(* IEC 61131-3 sources: Masterarbeit/sigmatek/lasalclass2/PW022_hardware/Class/SafetyManager (part 2) *)

          // if it has an active connection
          if pHelpManaging^.FlexCon.pFSoEConnection then
            // check if one of the safety number is the list match the one of the managing module
            pHelpHDINT := pPara^.aPara[1]$^HDINT;
            for i := 0 to (pPara^.aPara[0]-1)$UDINT do
              // if the connected number from the HWK is found in the list of connected numbers from the SCP => remember it to send it to the managing module
              if pHelpManaging^.FlexCon.SafetyNumber = pHelpHDINT^ then
                MyPara.aPara[0] := pHelpHDINT^$DINT;

                // stop searching for this managing device
                exit;
              end_if;

              pHelpHDINT += sizeof(HDINT);
            end_for;
          end_if;

          // send the current number for this device
          pHelpManaging^.pThis^.NewInst(#MyPara, #MyResult);

          pHelpManaging := pHelpManaging^.pNext;
        end_while;
      end_if;

//**********************************************************************************************************************************************************
    CMD_HWC_CONVERT_COMPRESSED_HWPATH:

      //Method is used to search through the configuration for the handed over compressed hw path and returns the respective uncompressed hw path

      //pPara^.aPara[0] .. version
      //pPara^.aPara[1] .. comp hw path
      //pPara^.aPara[2] .. comp hw path length
      //pPara^.aPara[3] .. pointer to buffer where hw path will be copied
      //pPara^.aPara[4] .. size of buffer where data will be copied

      //pResult^.aData[0]$DINT .. version
      //pResult^.aData[4]$DINT .. retcode when error (negative) or amount of bytes of hw path

      //Check for valid pointer and data lengths
      if (pPara^.aPara[1] = NIL)
       | (pPara^.aPara[2] = 0)
       | (pPara^.aPara[3] = NIL)
       | (pPara^.aPara[4] = 0) then

        ret_code := ERROR;
        pResult^.uiLng := 8;
        pResult^.aData[0]$DINT := 1;  //version of command
        pResult^.aData[4]$DINT := -1; //Invalid pointer or length
        return;
      end_if;

      if pConfigs = NIL  then
        ret_code := ERROR;
        pResult^.uiLng := 8;
        pResult^.aData[0]$DINT := 1;  //version of command
        pResult^.aData[4]$DINT := -2; //no configs yet
        return;
      end_if;

      pHelpConfigs := pConfigs;

      while pHelpConfigs do

        //Go through module configs
        //=============================================================================================================
        if pHelpConfigs^.pFirstModuleCfg then
          pHelpModuleConf := pHelpConfigs^.pFirstModuleCfg;

          while pHelpModuleConf do

            //Check if we got a valid path and len
            if pHelpModuleConf^.ModuleInfo.pCompPath & pHelpModuleConf^.ModuleInfo.CompPathLen then

              //Check if we found the passed path
              if _memcmp(ptr1:=pPara^.aPara[1]$^void, ptr2:=pHelpModuleConf^.ModuleInfo.pCompPath, cntr:=pPara^.aPara[2]$UDINT) = 0 then

                //we found the compressed hw path, return pointer to normal hw path
                if pPara^.aPara[4] > pHelpModuleConf^.ModuleInfo.PathLen then

                  //Copy path to user pointer
                  _memcpy(ptr1:=pPara^.aPara[3]$^void, ptr2:=pHelpModuleConf^.ModuleInfo.pPath, cntr:=pHelpModuleConf^.ModuleInfo.PathLen);

                  ret_code := READY;
                  pResult^.uiLng := 8;

                  pResult^.aData[0]$DINT := 1;  //version
                  pResult^.aData[4]$DINT := pHelpModuleConf^.ModuleInfo.PathLen;
                  return;

                else
                  ret_code := ERROR;
                  pResult^.uiLng := 8;
                  pResult^.aData[0]$DINT := 1;   //version
                  pResult^.aData[4]$DINT := -3;  //not enough space to copy path
                  return;

                end_if;

              end_if;
            end_if;
            pHelpModuleConf := pHelpModuleConf^.pNext;
          end_while;
        end_if;

        //Go through slave config
        //=============================================================================================================
        if pHelpConfigs^.pFirstSlaveCfg then

          pHelpSlaveCfg := pHelpConfigs^.pFirstSlaveCfg;

          while pHelpSlaveCfg do

            //Check if we got a valid path and len
            if pHelpSlaveCfg^.SlaveInfo.pCompPath & pHelpSlaveCfg^.SlaveInfo.CompPathLen then

              //Check if we found the passed path
              if _memcmp(ptr1:=pPara^.aPara[1]$^void, ptr2:=pHelpSlaveCfg^.SlaveInfo.pCompPath, cntr:=pPara^.aPara[2]$UDINT) = 0 then

                //we found the compressed hw path, return pointer to normal hw path
                if pPara^.aPara[4] > pHelpSlaveCfg^.SlaveInfo.PathLen then

                  //Copy path to user pointer
                  _memcpy(ptr1:=pPara^.aPara[3]$^void, ptr2:=pHelpSlaveCfg^.SlaveInfo.pPath, cntr:=pHelpSlaveCfg^.SlaveInfo.PathLen);

                  ret_code := READY;
                  pResult^.uiLng := 8;

                  pResult^.aData[0]$DINT := 1;  //Path was found
                  pResult^.aData[4]$DINT := pHelpSlaveCfg^.SlaveInfo.PathLen;
                  return;

                else
                  ret_code := ERROR;
                  pResult^.uiLng := 8;
                  pResult^.aData[0]$DINT := 1;   //version
                  pResult^.aData[4]$DINT := -3;  //not enough space to copy path
                  return;

                end_if;
              end_if;
            end_if;
            pHelpSlaveCfg := pHelpSlaveCfg^.pNext;
          end_while;
        end_if;

        //Go through fsoe connections
        //=============================================================================================================
        if pHelpConfigs^.pFirstFSoEConnection then
          pHelpFsoeConn := pHelpConfigs^.pFirstFSoEConnection;

          while pHelpFsoeConn do

            //Check if we got a valid path and len
            if pHelpFsoeConn^.pSlavePathComp & pHelpFsoeConn^.SlavePathLen then

              //Check if we found the passed path
              if _memcmp(ptr1:=pPara^.aPara[1]$^void, ptr2:=pHelpFsoeConn^.pSlavePathComp, cntr:=pPara^.aPara[2]$UDINT) = 0 then

                //we found the compressed hw path, return pointer to normal hw path
                if pPara^.aPara[4] > pHelpFsoeConn^.SlavePathLen then

                  //Copy path to user pointer
                  _memcpy(ptr1:=pPara^.aPara[3]$^void, ptr2:=pHelpFsoeConn^.pSlavePath, cntr:=pHelpFsoeConn^.SlavePathLen);

                  ret_code := READY;
                  pResult^.uiLng := 8;

                  pResult^.aData[0]$DINT := 1;  //Path was found
                  pResult^.aData[4]$DINT := pHelpFsoeConn^.SlavePathLen;
                  return;

                else
                  ret_code := ERROR;
                  pResult^.uiLng := 8;
                  pResult^.aData[0]$DINT := 1;   //version
                  pResult^.aData[4]$DINT := -3;  //not enough space to copy path
                  return;
                end_if;
              end_if;

            end_if;
            pHelpFsoeConn := pHelpFsoeConn^.pNext;
          end_while;
        end_if;

        pHelpConfigs := pHelpConfigs^.pNext;
      end_while;

      //comp hw path was not found in config
      ret_code := ERROR;
      pResult^.uiLng := 8;
      pResult^.aData[0]$DINT := 1;   //version
      pResult^.aData[4]$DINT := -4;  //passed path was not found in configuration list

//**********************************************************************************************************************************************************
  else
    bd_LogRtMessagesInCy.InvalidCommandReceived := TRUE;
  END_CASE;

#ifdef SAFETY_DEBUG_LOGGING_ACTIVATED
  if InitSSW <> OldInitSSW then
#ifdef SAFETY_DEBUG_TRACING_ACTIVATED
    LogValue("@DBG (SafetyManager::ClassState::NewInst) InitSSW changed from {0} to {1}", Value:=OldInitSSW, Value2:=InitSSW);
#endif
    LogBuf[ActLogIndex].NewState := InitSSW;
    LogBuf[ActLogIndex].OldState := OldInitSSW;
    LogBuf[ActLogIndex].Command := 0;
    LogBuf[ActLogIndex].TimeSinceLastLog_us := OS_READMICROSEC();
    LogBuf[ActLogIndex].TimeSinceLastLog_us -= TimeStampLastLog_us;
    TimeStampLastLog_us := OS_READMICROSEC();
    if ActLogIndex = (LogBufferSize - 1) then
      ActLogIndex := 0;
    else
      ActLogIndex += 1;
    end_if;
  end_if;
  OldInitSSW := InitSSW;
#endif

  ret_code := READY;

END_FUNCTION

FUNCTION VIRTUAL GLOBAL SafetyManager::CyWork
  VAR_INPUT
    EAX 	: UDINT;
  END_VAR
  VAR_OUTPUT
    state (EAX) 	: UDINT;
  END_VAR
  VAR
    MyPara 	      : CmdStruct;
    MyResult	    : results;
    pHelpSafety   : ^t_SafetyComponent;
    pHelpManaging : ^t_ManagingComponent;
    pModuleInfo   : ^t_ModuleInfo;
    pTempMem      : ^void;
    i             : UDINT;
    Synchron      : BOOL;
    AllReady      : BOOL;
    pHelpCfg      : ^t_LocalCfgListElem;
    pHelpConfig   : ^t_CfgListElem;
  END_VAR

//=================================================================================================
#ifdef VM_CLASS_TIME_MEASUREMENT
  StartTimeMeasurement(VARANTIME_CY);
#endif
//=================================================================================================
  // if we got UDP stuff going on => start the udp task
  if (sUdpVars.UdpTaskStarted = FALSE) & (sUdpVars.ProducerConnectionNo | ((sUdpVars.UdpInit AND 2#11) = (t_UdpInit.FSoEAvailable OR t_UdpInit.ProvidesIF))) then
    To_MultiTask.CREATETHREAD(taskfunction0 := #UdpTask()
                            , priority0     := 14           // same priority as cyclic task
                            , stackSize0    := 0x4000
                            , flags0        := MT_TASK_SAVETHIS
                            , parameter0    := THIS
                            , name0         := "SafetyUDP");

    sUdpVars.UdpTaskStarted := TRUE;
  end_if;

  case InitSSW of
//**********************************************************************************************************************************************************
    _NotMaster: // don't start any actions, because we're not the master. but if the master wants something from us, we help out

//**********************************************************************************************************************************************************
    _ClearRoutingInfos: // initialize the structures or clean up an old configuration
      if ClearRoutingInformations() then

        // reactivate the domain synchronicity timeout
        b_SynchroTimeoutSet := FALSE;

        InitSSW := _FirstWait4SynchronManagingNodes;
      end_if;

//**********************************************************************************************************************************************************
    _FirstWait4SynchronManagingNodes: // wait for managing nodes to be syncron (all nodes are optionaly for this case, the will be checked later again)
      if SafetyDomainTimeout & (b_SynchroTimeoutSet = FALSE) then
        b_SynchroTimeoutSet := TRUE;
        SynchroTimeout := ops.tAbsolute;
      end_if;

      Synchron := AllManagingNodesSynchron();
                                                        // we wait synchro timeout + 50ms (50ms time for the domains to give up trying: see AllManagingNodesSynchron method)
      if Synchron then// | (SafetyDomainTimeout & ((ops.tAbsolute - SynchroTimeout) > (SafetyDomainTimeout + 50))) then
        if b_SyncTimeoutExceeded then
          b_SyncTimeoutExceeded := FALSE;
          LogError("@0444 (SafetyManager::CyWork) Timeout for managing module (VBC, VMC,..) exceeded! Initialisation will continue to check if it's optional!");
        end_if;

        InitSSW := _SetConnectionOk;
      end_if;

//**********************************************************************************************************************************************************
    _SetConnectionOk:
      // send hw-connection ok to start SDOs
      MyPara.uiCmd := CMD_SM_FIRST_CONNECT_READY;
      MyPara.aPara[0] := 0; // length of parameters

      TellAllSafetyModules(#MyPara, #MyResult);

      b_MandatoryStuffAvailable := FALSE;
      LastCfgReceiveTime := ops.tAbsolute;

      InitSSW := _Wait4ReInit;

//**********************************************************************************************************************************************************
    _Wait4ReInit: // wait until all local CSCPs have a valid configuration before we wait to be synchron with other domains

      // add our local configurations if there are any
      SendLocalCfgsToMaster();

      // wait until we got a valid config of every local safety cpu
      if (LocalCPUCfgNo = LocalCPUNo) | b_MandatoryStuffAvailable then
        AllReady := TRUE;

        if LocalCPUCfgNo then
          pHelpCfg := pFirstLocalCPUCfg;

          // for is used to ensure thread safety
          for i := 0 to (LocalCPUCfgNo-1) do
            if pHelpCfg^.ConfigSize = 0 then
              AllReady := FALSE;
              exit;
            end_if;

            pHelpCfg := pHelpCfg^.pNext;
          end_for;
        end_if;

        // if we have a config from every cscp, we start the initialisation
        if AllReady then
          InitSSW := _CheckLocalCPUConfigs;
        end_if;
      else
        // if we already got a config => check if there is something optional
        if LocalCPUCfgNo & ((ops.tAbsolute - LastCfgReceiveTime) > 5000) then
          CheckOptional();
        end_if;

        InitSSW := _SendInterfaceConfigs;
      end_if;

//**********************************************************************************************************************************************************
    _CheckLocalCPUConfigs: // check for unused and optional modules in the local configurations (needed for correct time synchronisation)
      // if we have a configuration of every safety cpu => check if the managing modules are optional or any of the safety/managing components is unused (not involved in any PDO)
      if (LocalCPUCfgNo = LocalCPUNo) | b_MandatoryStuffAvailable then

        // set the IsOptional-Bit of all modules (safety and managing components) to TRUE
        // in CheckModuleUsage the the non-optional will get the IsOptional-Bit set to FALSE
        pHelpSafety := pFirstSafetyComponent;
        while pHelpSafety do
          pHelpSafety^.InfoBits.IsOptional    := TRUE;

          pHelpSafety := pHelpSafety^.pNext;
        end_while;

        pHelpManaging := pFirstManagingInterfaceComponent;
        while pHelpManaging do
          pHelpManaging^.InfoBits.IsOptional    := TRUE;

          pHelpManaging := pHelpManaging^.pNext;
        end_while;

        // check all configurations which modules are used
        if LocalCPUCfgNo then
          pHelpCfg := pFirstLocalCPUCfg;

          for i := 0 to (LocalCPUCfgNo-1) do
            // check for used modules and mark them in the infobits
            CheckModuleUsage(pHelpCfg^.ConfigSize, pHelpCfg^.pConfig, pHelpCfg^.IsFSoECfg);

            pHelpCfg := pHelpCfg^.pNext;
          end_for;
        end_if;

        // now create the linked list for the time synchronisation
        CreateTimeSyncList();

        if (pFirstManagingInterfaceComponent = NIL) then
          // if we have FSoE Modules => check the connection between the modules and tell them what to copy
          if b_GotFSoEModules then
            CreateFSoEPDOs();

            if b_AllLocalSlaveAddressesValid then
              InitSSW := _NoDomains;
            else
              // wait for all local connections to be established
              SetTimeout();
              InitSSW := _Wait4FSoEConnectionsLocal;
            end_if;
          else
            InitSSW := _NoDomains;
          end_if;
        else
          // reactivate the domain synchronicity timeout, because now we know what is really optional
          b_SynchroTimeoutSet := FALSE;

          InitSSW := _Wait4SynchronManagingNodes;
        end_if;

      end_if;

//**********************************************************************************************************************************************************
    _Wait4FSoEConnectionsLocal:
      CheckTimeout();
      if b_AllLocalSlaveAddressesValid then
        CreateFSoEPDOs();
        // success => continue
        InitSSW := _NoDomains;
      end_if;

//**********************************************************************************************************************************************************
    _Wait4SynchronManagingNodes: // wait until all managing modules are synchron with the other stations
      if SafetyDomainTimeout & (b_SynchroTimeoutSet = FALSE) then
        b_SynchroTimeoutSet := TRUE;
        SynchroTimeout := ops.tAbsolute;
      end_if;

      Synchron := AllManagingNodesSynchron();
                                                        // we wait synchro timeout + 50ms (50ms time for the domains to give up trying: see AllManagingNodesSynchron method)
      if Synchron then// | (SafetyDomainTimeout & ((ops.tAbsolute - SynchroTimeout) > (SafetyDomainTimeout + 50))) then
        if b_SyncTimeoutExceeded then
          b_SyncTimeoutExceeded := FALSE;
          LogError("@0445 (SafetyManager::CyWork) Timeout for optional managing module (VBC, VMC,..) exceeded! Initialisation will continue without it!");
        end_if;

        // add our own safety cpus to the config list
        AddOwnCPUsToList();

        if NewTimeSyncPossible() then
          // tell every safety module, that it has to initialize the memory for writing the time synchronisation
          SetNewSyncMode(TRUE);
          MyPara.aPara[3] := 1;
        else
          SetNewSyncMode(FALSE);
          MyPara.aPara[3] := 0;
        end_if;

        InitSSW := _SendDomainNr;
      end_if;

//**********************************************************************************************************************************************************
    _SendDomainNr: // send the domain nr. to the managing nodes
      // if we have a valid domain number
      MyPara.uiCmd := CMD_SM_DOMAIN_NR_SEND;
      MyPara.aPara[0] := 1; // length of parameters

      pTempMem := NIL;

      if us_SafetyModuleNo then
        if ud_SizeTempMemCy >= 1 + us_SafetyModuleNo * sizeof(t_ModuleInfo) then
          pTempMem := pTempMemCy;
        else
          LogError("@0446 (SafetyManager::CyWork) _SendDomainNr: Temporary memory for cyclic task is too small!");
          LogValue("AvaliableMem: {0} / NeededMem: {1}", Value:=ud_SizeTempMemCy, Value2:=1 + us_SafetyModuleNo * sizeof(t_ModuleInfo));
        end_if;

        if pTempMem then
          MyPara.aPara[1] := pTempMem$DINT;
          pModuleInfo$^void := pTempMem;

          pModuleInfo^$USINT := 0;
          pModuleInfo += sizeof(USINT);
          if pFirstSafetyComponent then
            pHelpSafety := pFirstSafetyComponent;
            while pHelpSafety do
              pModuleInfo^.SafetyNbr := pHelpSafety^.SafetyNbr;

              pHelpSafety := pHelpSafety^.pNext;
              pModuleInfo += sizeof(t_ModuleInfo);
            end_while;

            MyPara.aPara[0] += us_SafetyModuleNo * sizeof(t_ModuleInfo);
          end_if;
        else
          MyPara.aPara[1] := (#MyPara.aPara[3])$DINT;
          MyPara.aPara[3] := 0;
          LogError("@0447 (SafetyManager::CyWork) Failed to allocate memory for distributing the local module information");
        end_if;
      else
        MyPara.aPara[1] := (#MyPara.aPara[3])$DINT;
        MyPara.aPara[3] := 0;
      end_if;

      // tell all interface modules, because maybe they don't know we're an interface neighbor
      TellAllInterfaceManagingModules(#MyPara, #MyResult);

      DomainInfoSendTime := ops.tAbsolute;

      // the slaves get this via newinst command
      InitSSW := _Wait4DomainInfos;

//**********************************************************************************************************************************************************
    _Wait4DomainInfos:
      // wait a little for further domain infos (which are sent as response to our message)
      if (ops.tAbsolute - DomainInfoSendTime) > 200 then
        InitSSW := _Wait4CPUConfigs;
        SetTimeout();
      end_if;

//**********************************************************************************************************************************************************
    _Wait4CPUConfigs:
      CheckTimeout();
      if AllCPUConfigsArrived() then
        // if all needed modules are available (all non-optional modules or interface frames)
        if CheckCPUConfigs() then
          // check if there are PDO configs to broadcast
          if ActPDO_ID then
            // before we broadcast the PDOs, we check if the length informations are correct on every entry
            PDOLengthCorrection();

            // if we have interface-connections, we wait for the safety numbers of it
            if pFirstManagingInterfaceComponent & AnyIFDomainSynchron() then
              InitSSW := _SendInterfaceConfigs;
            else
              InitSSW := _SendNextPDO;
            end_if;
          else
            if pFirstManagingInterfaceComponent & b_GotFSoEModules then
              // we have some FSoE Connections
              InitSSW := _SendInterfaceConfigs;
            else
              // otherwise => finalize initialisation
              InitSSW := _Wait4CopyCmdStart;
            end_if;
          end_if;
        else
          // if configs are not ok => set everything to finished so that the firmware can show the error information (otherwise the firmware will not start doing anything)
          InitSSW := _Wait4CopyCmdStart;
        end_if;
      end_if;

//**********************************************************************************************************************************************************
    _SendInterfaceConfigs:
      // if all domain managing modules needed for non-optional pdos are synchron
      if AllNonOptionalIFDomainsSynchron() then
        if b_GotFSoEModules then
          CreateFSoEPDOs();
        end_if;

        // send our configs to all inferface domains
        SendInterfaceConfigs(NIL, FALSE, b_GotFSoEModules);

        InitSSW := _Wait4InterfaceConfigs;
        SetTimeout();
      end_if;

//**********************************************************************************************************************************************************
    _Wait4InterfaceConfigs:
      CheckTimeout();
      if AllInterfaceCfgsArrived() then
        if (LocalCPUCfgNo = LocalCPUNo) | b_MandatoryStuffAvailable then
          if pActualSendPDO then
            InitSSW := _SendNextPDO;
          else
            if b_GotFSoEModules then
              SetTimeout();
              InitSSW := _Wait4FSoEConnectionsExternal;
            else
              InitSSW := _Wait4ReInit;
            end_if;
          end_if;
        else
          InitSSW := _Wait4ReInit;
        end_If;
      end_if;

//**********************************************************************************************************************************************************
    _Wait4FSoEConnectionsExternal:
      CheckTimeout();
      if b_AllLocalSlaveAddressesValid then
        CreateFSoEPDOs();
        FinalizePDOMapping();
        InitSSW := _FinishInitialisation;
      end_if;

//**********************************************************************************************************************************************************
    _SendNextPDO:
      // broadcast the PDO
      BroadCastActPDO();

      InitSSW := _Wait4PDOAcks;
      SetTimeout();

//**********************************************************************************************************************************************************
    _Wait4PDOAcks:
      // wait until all acknowledges arrive (all modules which are needed for PDO transport have to answer!)
      CheckTimeout();

      // check if there is another PDO configuration to send
      repeat
        if pActualSendPDO^.pNext then
          pActualSendPDO := pActualSendPDO^.pNext;
        else
          if pActualSendCfg^.pNext then
            pActualSendCfg := pActualSendCfg^.pNext;
            pActualSendPDO := pActualSendCfg^.pFirstPdoCfg;

            // if there is no pdo config in this config, go to the next config
            while (pActualSendPDO = NIL) & pActualSendCfg^.pNext do
              pActualSendCfg := pActualSendCfg^.pNext;
              pActualSendPDO := pActualSendCfg^.pFirstPdoCfg;
            end_while;
          else
            pActualSendCfg := NIL;
            pActualSendPDO := NIL;
          end_if;
        end_if;

      // skip double entries
      until ((pActualSendPDO = NIL) | (pActualSendPDO^.PdoInfo.Info.DoublePDOEntry = FALSE)) end_repeat;

      // if we found another PDO => send it
      if pActualSendPDO then
        InitSSW := _SendNextPDO;
      else
        // otherwise => finalize initialisation
        InitSSW := _Wait4CopyCmdStart;
      end_if;

//**********************************************************************************************************************************************************
    _Wait4CopyCmdStart:
      // this step is handlet in RT because the DOs are isochronous

//**********************************************************************************************************************************************************
    _NoDomains:
      // No domains available => just check if there are old modules or new modules used
      if NewTimeSyncPossible() then
        // tell every safety module, that it has to initialize the memory for writing the time synchronisation
        SetNewSyncMode(TRUE);
      else
        SetNewSyncMode(FALSE);
      end_if;

      // we may have internal interface frames and therefore we have to create a list with the local CRCs
      if LocalIFsAvailable() then
        // add local IFs for easier SDO/TDO forwarding
        CheckCPUConfigs();

        // check if there are PDO configs to broadcast
        if ActPDO_ID & (b_GotFSoEModules = FALSE) then
          // before we broadcast the PDOs, we check if the length informations are correct on every entry
          PDOLengthCorrection();

          // distribute PDOs locally
          pHelpConfig := pConfigs;
          while pHelpConfig do
            pActualSendCfg := pHelpConfig;
            pActualSendPDO := pHelpConfig^.pFirstPdoCfg;
            while pActualSendPDO do
              BroadCastActPDO();

              pActualSendPDO := pActualSendPDO^.pNext;
            end_while;

            pHelpConfig := pHelpConfig^.pNext;
          end_while;
        end_if;
      end_if;

      InitSSW := _FinishInitialisation;

//**********************************************************************************************************************************************************
    _FinishInitialisation:
      // if it's the new mode also start the sync process at the first safety device
      MyPara.uiCmd := CMD_SM_INIT_FINISHED;
      MyPara.aPara[0] := 0; // length of parameters

      // sent set bus ready signal (quit error 199 if active)
      TellAllSafetyModules(#MyPara, #MyResult);

      // if we have the new sync mode => start the time synchronisation here
      if b_NewSyncMode then
        b_StartTimeSync := TRUE;
      end_if;

      MinSyncDuration := 16#7FFFFFFF;

      // if there was an error and we still reached this point, don't conceal the error (except if it's a timeout in this init sequence or a SDO problem which could have been fixed)
      if (ClassState = 0) | (ClassState = -11) | (ClassState = -8) then
        ClassState := 1;
      end_if;

      InitSSW := _InitFinished;

//**********************************************************************************************************************************************************
    _InitFinished: // finished with initialisation, now start our cyclic business

      // check sync timeout counter
      if SyncTimeoutCounter >= TIMESYNC_TIMEOUTS_BEFORE_LOGMSG then
        LogError("@0448 (SafetyManager::CyWork) Timeout while Timesynchronizing");

        // reset counter
        SyncTimeoutCounter := 0;
      end_if;

      // print log messages from realtime here to prevent rt-runtime errors
      if bd_LogRtMessagesInCy then
        if bd_LogRtMessagesInCy.NoTDOTargetToManager then
          bd_LogRtMessagesInCy.NoTDOTargetToManager := FALSE;
          LogError("@0449 (SafetyManager::ClassState::NewInst) Couldn't find target of TDO on the way to the manager");
        end_if;

        if bd_LogRtMessagesInCy.NoTDOTargetToModule then
          bd_LogRtMessagesInCy.NoTDOTargetToModule := FALSE;
          LogError("@044A (SafetyManager::ClassState::NewInst) Couldn't find target of TDO on the way to the module");
        end_if;

        if bd_LogRtMessagesInCy.InvalidCommandReceived then
          bd_LogRtMessagesInCy.InvalidCommandReceived := FALSE;
          LogError("@044B (SafetyManager::State::NewInst) Invalid command received");
        end_if;

        if bd_LogRtMessagesInCy.UnkownCopySource then
          bd_LogRtMessagesInCy.UnkownCopySource := FALSE;
          LogError("@044D (SafetyManager::RtWork) Could not activate copy command, because source address is unknown (waiting for safety number info)");
        end_if;

        if bd_LogRtMessagesInCy.InvalidIFConfiguration then
          bd_LogRtMessagesInCy.InvalidIFConfiguration := FALSE;
          LogError("@044E (SafetyManager::GiveTokenToNextModule) Only non-synchron interface domains found => need at least one safe CPU!");
        end_if;

        if bd_LogRtMessagesInCy.TooManyOptionalMissing then
          bd_LogRtMessagesInCy.TooManyOptionalMissing := FALSE;
          LogError("@044F (SafetyManager::GiveTokenToNextModule) Too many optional modules missing for a correct time sync cycle");
        end_if;

        if bd_LogRtMessagesInCy.UdpReceivedInvalidCommand then
          bd_LogRtMessagesInCy.UdpReceivedInvalidCommand := FALSE;
          LogError("@0450 (SafetyManager::ReceiveUdpData) Received invalid command via UDP");
        end_if;

        if bd_LogRtMessagesInCy.UdpReceivedInvalidState then
          bd_LogRtMessagesInCy.UdpReceivedInvalidState := FALSE;
          LogError("@0451 (SafetyManager::ReceiveUdpData) Received invalid state via UDP");
        end_if;

        if bd_LogRtMessagesInCy.UdpNoMem4Connections then
          bd_LogRtMessagesInCy.UdpNoMem4Connections := FALSE;
          LogError("@0452 (SafetyManager::AddIpConnection) Can't add udp connection, since the memory is not allocated");
        end_if;
      end_if;
//**********************************************************************************************************************************************************
  end_case;

#ifdef SAFETY_DEBUG_LOGGING_ACTIVATED
  if InitSSW <> OldInitSSW then
#ifdef SAFETY_DEBUG_TRACING_ACTIVATED
    LogValue("@DBG (SafetyManager::CyWork) InitSSW changed from {0} to {1}", Value:=OldInitSSW, Value2:=InitSSW);
#endif
    LogBuf[ActLogIndex].NewState := InitSSW;
    LogBuf[ActLogIndex].OldState := OldInitSSW;
    LogBuf[ActLogIndex].Command := 0;
    LogBuf[ActLogIndex].TimeSinceLastLog_us := OS_READMICROSEC();
    LogBuf[ActLogIndex].TimeSinceLastLog_us -= TimeStampLastLog_us;
    TimeStampLastLog_us := OS_READMICROSEC();
    if ActLogIndex = (LogBufferSize - 1) then
      ActLogIndex := 0;
    else
      ActLogIndex += 1;
    end_if;
  end_if;
  OldInitSSW := InitSSW;
#endif

  state := READY;

//=================================================================================================
#ifdef VM_CLASS_TIME_MEASUREMENT
  StopTimeMeasurement(VARANTIME_CY);
#endif
//=================================================================================================

END_FUNCTION

FUNCTION SafetyManager::AddModule
  VAR_INPUT
    pPara 	: ^CmdStruct;
  END_VAR
  VAR_OUTPUT
    retcode 	: BOOL;
  END_VAR
  VAR
    ModuleType : t_e_ModuleType;
  END_VAR

  retcode := FALSE;

  ModuleType := pPara^.aPara[0]$t_e_ModuleType;

  // we differ between real safety components and managing components
  case ModuleType of
    _CSCP01x,
    _CSDI16x,
    _CSTO08x,
    _SCP010,
    _SCP011,
    _SCP111,
    _SCP211,
    _MS011,
    _MS012,
    _SDD1300,
    _SDD1400,
    _SDD1500,
    _SDD1600,
    _ModuleWithoutConfig:
        retcode := AddSafetyModule(ModuleType, pPara^.aPara[1]$pVirtualBase);

        if IsFSoEModule(ModuleType) then

          //only allocate memory if it is not done before
          if sUdpVars.pTempSendBufferCy = NIL then
            // allocate memory for the temporary cyclic send buffer
            sUdpVars.pTempSendBufferCy$pVoid := To_StdLib.Malloc(size:=sizeof(t_UdpPacketV2));

            if sUdpVars.pTempSendBufferCy then
              _memset(dest:=sUdpVars.pTempSendBufferCy, usByte:=0, cntr:=sizeof(t_UdpPacketV2));
            else
              SetError(bError:=TRUE, ErrorMessage:=_NO_MEMORY_SENDBUFFER_UDP_ERROR, dError:=0);
              LogError("@0453 (SafetyManager::AddModule) Failed to allocate memory for udp send buffer");
            end_if;
          end_if;

          //only allocate memory if it is not done before
          if sUdpVars.pTempSendBufferIRQ = NIL then
            // allocate memory for the temporary irq send buffer
            sUdpVars.pTempSendBufferIRQ$pVoid := To_StdLib.Malloc(size:=sizeof(t_UdpPacketV2));

            if sUdpVars.pTempSendBufferIRQ then
              _memset(dest:=sUdpVars.pTempSendBufferIRQ, usByte:=0, cntr:=sizeof(t_UdpPacketV2));
            else
              SetError(bError:=TRUE, ErrorMessage:=_NO_MEMORY_SENDBUFFER_UDP_ERROR, dError:=0);
              LogError("@0453 (SafetyManager::AddModule) Failed to allocate memory for udp send buffer");
            end_if;
          end_if;

          //only allocate memory if it is not done before
          if sUdpVars.paConnectionsToProducers = NIL then
            sUdpVars.paConnectionsToProducers$pVoid := To_StdLib.Malloc(size:=sizeof(t_aUdpConnections));

            if sUdpVars.paConnectionsToProducers then
              _memset(dest:=sUdpVars.paConnectionsToProducers, usByte:=0, cntr:=sizeof(t_aUdpConnections));
            else
              SetError(bError:=TRUE, ErrorMessage:=_NO_MEMORY_CONNECTION_BUFFER_UDP_ERROR, dError:=0);
              LogError("@0454 (SafetyManager::AddModule) Failed to allocate memory for udp receive buffer");
            end_if;
          end_if;

          //only allocate memory if it is not done before
          if sUdpVars.paConnectionsToConsumers = NIL then
            sUdpVars.paConnectionsToConsumers$pVoid := To_StdLib.Malloc(size:=sizeof(t_aUdpConnections));

            if sUdpVars.paConnectionsToConsumers then
              _memset(dest:=sUdpVars.paConnectionsToConsumers, usByte:=0, cntr:=sizeof(t_aUdpConnections));
            else
              SetError(bError:=TRUE, ErrorMessage:=_NO_MEMORY_CONNECTION_BUFFER_UDP_ERROR, dError:=0);
              LogError("@0454 (SafetyManager::AddModule) Failed to allocate memory for udp receive buffer");
            end_if;
          end_if;
        end_if;

    _VBC021Master,
    _VBC021Slave, // (is limited to 1 per system, because the system can't sync to different systems at the same time)
    _VMC052,
    _VaranManager4VMC, // VaranManager (VMC052 counterpart is also limited to 1 per system, because the system can't sync to different systems at the same time)
    _GenericTimeSyncMaster,
    _GenericTimeSyncSlave,
    _GenericFSoE:
        retcode := AddManagingModule(ModuleType, pPara^.aPara[1]$pVirtualBase, pPara^.aPara[2]$^USINT);
    _GenericDynamicFSoE:
        retcode := AddGenericDynamic(ModuleType, pPara^.aPara[1]$pVirtualBase, pPara^.aPara[2]$^USINT);
  else
    // invalid module type
    ClassState := -7;
    LogError("@0455 (SafetyManager::AddModule) Invalid ModuleType");
  end_case;

  if retcode then
    LoginCnt += 1;
  end_if;

END_FUNCTION

FUNCTION SafetyManager::AddSafetyModule
  VAR_INPUT
    ModuleType 	: t_e_ModuleType;
    pThis 	: pVirtualBase;
  END_VAR
  VAR_OUTPUT
    retcode 	: BOOL;
  END_VAR
  VAR
    pHelpSafety : ^t_SafetyComponent;
  END_VAR

  if pFirstSafetyComponent = NIL then
    pFirstSafetyComponent$pVoid := To_StdLib.Malloc(size:=sizeof(t_SafetyComponent));
    pHelpSafety := pFirstSafetyComponent;
  else
    pHelpSafety := pFirstSafetyComponent;
    while pHelpSafety^.pNext <> NIL do
      pHelpSafety := pHelpSafety^.pNext;
    end_while;
    pHelpSafety^.pNext$pVoid := To_StdLib.Malloc(size:=sizeof(t_SafetyComponent));
    pHelpSafety := pHelpSafety^.pNext;
  end_if;

  if pHelpSafety <> NIL then
    _memset(dest:=pHelpSafety, usByte:=0, cntr:=sizeof(t_SafetyComponent));
    pHelpSafety^.ModuleType   := ModuleType;
    pHelpSafety^.pThis        := pThis;

//    pHelpSafety^.pNext        := NIL;  // not necessary because of memset

    case ModuleType of
//**********************************************************************************************************************************************************
      _CSCP01x,
      _SCP010,
      _SCP011,
      _SCP111,
      _SCP211,
      _SDD1300,
      _SDD1400,
      _SDD1500,
      _SDD1600:
        LocalCPUNo += 1;

//**********************************************************************************************************************************************************
      _CSDI16x,
      _MS011,
      _MS012:
        pHelpSafety^.InfoBits.OnlyInputs := TRUE;
//**********************************************************************************************************************************************************
    end_case;

    us_SafetyModuleNo += 1;

    retcode := TRUE;
  else
    ClassState := -1;

    retcode := FALSE;
  end_if;

END_FUNCTION

FUNCTION SafetyManager::AddManagingModule
  VAR_INPUT
    ModuleType 	: t_e_ModuleType;
    pThis 	: pVirtualBase;
    pObjectPath 	: ^USINT;
  END_VAR
  VAR_OUTPUT
    retcode 	: BOOL;
  END_VAR
  VAR
    pHelpManaging : ^t_ManagingComponent;
    pMyPath : ^USINT;
  END_VAR

  if pFirstManagingInterfaceComponent = NIL then
    pFirstManagingInterfaceComponent$pVoid := To_StdLib.Malloc(size:=sizeof(t_ManagingComponent));
    pHelpManaging := pFirstManagingInterfaceComponent;
  else
    pHelpManaging := pFirstManagingInterfaceComponent;
    while pHelpManaging^.pNext <> NIL do
      pHelpManaging := pHelpManaging^.pNext;
    end_while;
    pHelpManaging^.pNext$pVoid := To_StdLib.Malloc(size:=sizeof(t_ManagingComponent));
    pHelpManaging := pHelpManaging^.pNext;
  end_if;

  if pHelpManaging <> NIL then
    _memset(dest:=pHelpManaging, usByte:=0, cntr:=sizeof(t_ManagingComponent));
    pHelpManaging^.ModuleType     := ModuleType;
    pHelpManaging^.pThis          := pThis;
    pHelpManaging^.DomainNr       := 16#FF;

    if pObjectPath then
      pMyPath$^void := To_StdLib.Malloc(size:=pObjectPath^ + 2);

      // convert 1 byte length info into 2 byte length info
      if pMyPath then
        pMyPath^$UINT := pObjectPath^$USINT;
        To_StdLib.MemCpy(dest:=pMyPath + 2, source:=pObjectPath + 1, size:=pObjectPath^);
      end_if;
    end_if;

    pHelpManaging^.pModulePath := pMyPath;

  //pHelpManaging^.pNext          := NIL;  // not necessary because of memset

    retcode := TRUE;
  else
    ClassState := -1;

    retcode := FALSE;
  end_if;

END_FUNCTION

FUNCTION SafetyManager::AddGenericDynamic
  VAR_INPUT
    ModuleType 	: t_e_ModuleType;
    pThis 	: pVirtualBase;
    pObjectPath 	: ^USINT;
  END_VAR
  VAR_OUTPUT
    retcode 	: BOOL;
  END_VAR
  VAR
    pHelpManaging : ^t_GenericDynamicComponent;
    pMyPath : ^USINT;
  END_VAR

  if pFirstGenericDynamic = NIL then
    pFirstGenericDynamic$pVoid := To_StdLib.Malloc(size:=sizeof(t_GenericDynamicComponent));
    pHelpManaging := pFirstGenericDynamic;
  else
    pHelpManaging := pFirstGenericDynamic;
    while pHelpManaging^.pNext <> NIL do
      pHelpManaging := pHelpManaging^.pNext;
    end_while;
    pHelpManaging^.pNext$pVoid := To_StdLib.Malloc(size:=sizeof(t_GenericDynamicComponent));
    pHelpManaging := pHelpManaging^.pNext;
  end_if;

  if pHelpManaging <> NIL then
    _memset(dest:=pHelpManaging, usByte:=0, cntr:=sizeof(t_GenericDynamicComponent));
    pHelpManaging^.ModuleType     := ModuleType;
    pHelpManaging^.pThis          := pThis;

    if pObjectPath then
      pMyPath$^void := To_StdLib.Malloc(size:=pObjectPath^ + 2);

      // convert 1 byte length info into 2 byte length info
      if pMyPath then
        pMyPath^$UINT := pObjectPath^$USINT;
        To_StdLib.MemCpy(dest:=pMyPath + 2, source:=pObjectPath + 1, size:=pObjectPath^);
      end_if;
    end_if;

    pHelpManaging^.pModulePath := pMyPath;

  //pHelpManaging^.pNext          := NIL;  // not necessary because of memset

    retcode := TRUE;
  else
    ClassState := -1;

    retcode := FALSE;
  end_if;

END_FUNCTION

FUNCTION SafetyManager::AddSafetyNbr
	VAR_INPUT
		pThis 	: pVirtualBase;
		ud_SafetyNbr 	: HDINT;
		FirmwareVersion 	: HDINT;
		FPGAVersion 	: HSINT;
		PathLen 	: USINT;
		pPath 	: ^USINT;
	END_VAR
	VAR_OUTPUT
		retcode 	: BOOL;
	END_VAR
  VAR
    pHelpSafety             : ^t_SafetyComponent;
    pHelpConfigManager      : ^t_CfgListElem;
    pHelpConnectionManager  : ^t_FSoEConnectionDetails;
    pHelpModuleCfg          : ^t_ModuleListElem;
    MyPara 	                : CmdStruct;
    MyResult	              : results;
    pOwnerSafety            : ^t_SafetyComponent;
  END_VAR

  retcode := FALSE;

  if pFirstSafetyComponent then
    pHelpSafety := pFirstSafetyComponent;
    while pHelpSafety do
      if pHelpSafety^.pThis = pThis then
        pHelpSafety^.SafetyNbr    := ud_SafetyNbr;
        pHelpSafety^.FW_Version   := FirmwareVersion;
        pHelpSafety^.FPGA_Version := FPGAVersion;
        pHelpSafety^.PathLen      := PathLen;
        pHelpSafety^.pPath        := pPath;

        if pHelpSafety^.ModuleType = _ModuleWithoutConfig then

          // if the post init is finished => module added during runtime
          if b_PostInitFinished then

            // check all configs
            pHelpConfigManager := pConfigs;
            while pHelpConfigManager do

              // check for FSoE connections that haven't been initialized
              pHelpConnectionManager := pHelpConfigManager^.pFirstFSoEConnection;
              while pHelpConnectionManager do

                if pHelpConnectionManager^.Flags.FSoESlaveHasNoConfig & pHelpConnectionManager^.Flags.IsMaster then
                  if pHelpConnectionManager^.InternalConnectionState = FCS_RESET then
                    ShareSingleConnectionInfos(pHelpConnectionManager, pHelpConfigManager^.pFirstModuleCfg);
                  end_if;
                end_if;

                pHelpConnectionManager := pHelpConnectionManager^.pNext;
              end_while;

              // check all module configs for a match of the path and inform the owner that there is a new safety number
              pHelpModuleCfg := pHelpConfigManager^.pFirstModuleCfg;
              while pHelpModuleCfg do
                if (pHelpModuleCfg^.ModuleInfo.pPath^ = pPath^) &
                   (To_StdLib.MemCmp(pPath + 1, pHelpModuleCfg^.ModuleInfo.pPath + 2 + pHelpModuleCfg^.ModuleInfo.pPath^ - pPath^, pPath^) = 0) then

                  // found a match => tell the owner of the configuration we found the module in

                  pOwnerSafety := pFirstSafetyComponent;
                  while pOwnerSafety do
                    if pOwnerSafety^.SafetyNbr = pHelpConfigManager^.SafetyNbr then
                      MyPara.uiCmd    := CMD_SM_UPDATE_SAFETY_NBR;
                      MyPara.aPara[0] := pHelpModuleCfg^.ModuleInfo.CompPathLen;    // length of HW path
                      MyPara.aPara[1] := pHelpModuleCfg^.ModuleInfo.pCompPath$DINT; // pointer to HW path
                      MyPara.aPara[2] := ud_SafetyNbr$DINT;                         // new safety number
                      pOwnerSafety^.pThis^.NewInst(#MyPara, #MyResult);
                    end_if;

                    pOwnerSafety := pOwnerSafety^.pNext;
                  end_while;
                end_if;

                pHelpModuleCfg := pHelpModuleCfg^.pNext;
              end_while;

              pHelpConfigManager := pHelpConfigManager^.pNext;
            end_while;
          end_if;
        end_if;

        retcode := TRUE;
        return;
      end_if;

      pHelpSafety := pHelpSafety^.pNext;
    end_while;
  end_if;

END_FUNCTION

FUNCTION SafetyManager::GetModuleTypeNo
  VAR_INPUT
    ModuleType 	: t_e_ModuleType;
  END_VAR
  VAR_OUTPUT
    ModuleNo 	: UDINT;
  END_VAR
  VAR
    pHelpSafety   : ^t_SafetyComponent;
    pHelpManaging : ^t_ManagingComponent;
    pHelpGeneric        : ^t_GenericDynamicComponent;
  END_VAR

  ModuleNo := 0;

  if pFirstSafetyComponent then
    pHelpSafety := pFirstSafetyComponent;
    while pHelpSafety do
      if pHelpSafety^.ModuleType = ModuleType then
        ModuleNo += 1;
      end_if;

      pHelpSafety := pHelpSafety^.pNext;
    end_while;
  end_if;

  if pFirstManagingInterfaceComponent then
    pHelpManaging := pFirstManagingInterfaceComponent;
    while pHelpManaging do
      if pHelpManaging^.ModuleType = ModuleType then
        ModuleNo += 1;
      end_if;

      pHelpManaging := pHelpManaging^.pNext;
    end_while;
  end_if;

  if pFirstGenericDynamic then
    pHelpGeneric := pFirstGenericDynamic;

    while pHelpGeneric do
      if pHelpGeneric^.ModuleType = ModuleType then
        ModuleNo += 1;
      end_if;

      pHelpGeneric := pHelpGeneric^.pNext;
    end_while;

  end_if;

END_FUNCTION

FUNCTION SafetyManager::NewTimeSyncPossible
  VAR_OUTPUT
    retcode 	: BOOL;
  END_VAR
  VAR
    pHelpSafety   : ^t_SafetyComponent;
  END_VAR

  // if there is FSoE in the project => no timesync
  if b_GotFSoEModules then
    retcode := FALSE;
    return;
  end_if;

  // default is: we can => check if there is any module with too old firmware or fpga
  retcode := TRUE;

  if pFirstSafetyComponent then
    pHelpSafety := pFirstSafetyComponent;
    while pHelpSafety do

      // check all modules for correct versions
      if ((pHelpSafety^.ModuleType = _CSCP01x) & (   (pHelpSafety^.FPGA_Version    < 16#14)     // if its a CSCP and the FPGA Version is lower than 1.4
                                                   | (pHelpSafety^.FW_Version$UINT < 100)) &    // or the firmware version is lower than 100
                                                      pHelpSafety^.SafetyNbr)                   // only if there is a safety number available (maybe the module is optional and not available)
      |  (pHelpSafety^.NewConfigType = ConfigState_Old) then                                    // or the module has an old config type

        retcode := FALSE;
      end_if;

      pHelpSafety := pHelpSafety^.pNext;
    end_while;
  end_if;

END_FUNCTION

FUNCTION SafetyManager::SetNewSyncMode
  VAR_INPUT
    b_NewMode 	: BOOL;
  END_VAR
  VAR
    MyPara 	  : CmdStruct;
    MyResult	: results;
  END_VAR

  b_NewSyncMode := b_NewMode;

  MyPara.uiCmd := CMD_SM_SET_NEW_SYNC_MODE;
  MyPara.aPara[0] := b_NewSyncMode;
  TellAllSafetyModules(#MyPara, #MyResult);

END_FUNCTION

FUNCTION SafetyManager::TellAllSafetyModules
  VAR_INPUT
    pPara 	: ^CmdStruct;
    pResult 	: ^results;
  END_VAR
  VAR
    pHelpSafety : ^t_SafetyComponent;
  END_VAR

  if pFirstSafetyComponent then
    pHelpSafety := pFirstSafetyComponent;
    while pHelpSafety do
      // call the newinst with the given parameters
      pHelpSafety^.pThis^.NewInst(pPara, pResult);

      pHelpSafety := pHelpSafety^.pNext;
    end_while;
  end_if;

END_FUNCTION

FUNCTION SafetyManager::StartTimeSync

  if pFirstTimeSyncElement then
    pActTimeSyncElement := pFirstTimeSyncElement;

    // send the token to the right module
    GiveTokenToNextModule();

    // remember the start time for calculating the time of a complete synchronisation
    TimeSyncCycleStart := ops.tAbsolute;
  end_if;

END_FUNCTION

FUNCTION SafetyManager::NextTimeSyncModule

  pActTimeSyncElement := pActTimeSyncElement^.pNext;

  // must be done after selecting the new element
  if GiveTokenToNextModule() then
    // we're finished with our synchronisation cycle and just started a new one (must be done after selecting the new element)
    if IsTimeSyncMaster then
      SyncDuration := ops.tAbsolute - TimeSyncCycleStart;
      if SyncDuration > MaxSyncDuration then
        MaxSyncDuration := SyncDuration;
      end_if;
      if SyncDuration < MinSyncDuration then
        MinSyncDuration := SyncDuration;
      end_if;

      // if a cycle has been finished => reset the timeout counter
      SyncTimeoutCounter := 0;

      // remember the start time for calculating the time of a complete synchronisation
      TimeSyncCycleStart := ops.tAbsolute;
    end_if;
  end_if;

END_FUNCTION

FUNCTION SafetyManager::GiveTokenToNextModule
  VAR_OUTPUT
    RestartCycle 	: BOOL;
  END_VAR
  VAR
    MyPara 	  : CmdStruct;
    MyResult	: results;
    pTemp : ^t_TimeSyncElement;
  END_VAR

  if pActTimeSyncElement = pFirstTimeSyncElement then
    RestartCycle := TRUE;
  else
    RestartCycle := FALSE;
  end_if;

  // check if we have to skip something (missing optional modules)
  if TimeSyncModuleAvailable(pActTimeSyncElement) = FALSE then
    // save the actual position
    pTemp := pActTimeSyncElement;

    // if it's a missing optional module
    while (TimeSyncModuleAvailable(pActTimeSyncElement) = FALSE) do
      // skip it
      pActTimeSyncElement := pActTimeSyncElement^.pNext;

      // if we jumped on the first, we have to restart the cycle (time measurement and timeout surveillance)
      if pActTimeSyncElement = pFirstTimeSyncElement then
        RestartCycle := TRUE;
      end_if;

      // if we're at the start of the rotation => stop rotating and print error message
      if pActTimeSyncElement = pTemp then
        bd_LogRtMessagesInCy.TooManyOptionalMissing := TRUE;
        ClassState := -12;
        exit;
      end_if;
    end_while;
  end_if;

  // check if we have to skip something
  if pActTimeSyncElement^.InfoBits.IsInterfaceDomain then
    // save the actual position
    pTemp := pActTimeSyncElement;

    // if it's an interface managing module and it's not synchron, skip it (there has to be also a Safety CPU in the system, therefore we don't ask for it
    while pActTimeSyncElement^.InfoBits.IsInterfaceDomain & (pActTimeSyncElement^.pManaging^.InfoBits.IsSynchron = FALSE) do
      // skip it
      pActTimeSyncElement := pActTimeSyncElement^.pNext;

      // if we jumped on the first, we have to restart the cycle (time measurement and timeout surveillance)
      if pActTimeSyncElement = pFirstTimeSyncElement then
        RestartCycle := TRUE;
      end_if;

      // if we're at the start of the rotation => stop rotating and print error message
      if pActTimeSyncElement = pTemp then
        bd_LogRtMessagesInCy.InvalidIFConfiguration := TRUE;
        ClassState := -12;
        exit;
      end_if;
    end_while;
  end_if;

  if pActTimeSyncElement^.InfoBits.IsConnectionToMaster then
    // don't check for sync timeout if we're not the master
    b_CheckTimeSyncTimeout := FALSE;
  else
    b_CheckTimeSyncTimeout := TRUE;
  end_if;

  // if it's a managing module and not the connection to the master, we give the token to a slave => remember it
  if pActTimeSyncElement^.InfoBits.IsManagingModule & (pActTimeSyncElement^.InfoBits.IsConnectionToMaster = FALSE) then
    b_SlaveSyncActive := TRUE;
  end_if;

  // tell the next module, to start the time synchronisation
  MyPara.uiCmd := CMD_SM_START_TIME_SYNC;
  pActTimeSyncElement^.pThis^.NewInst(#MyPara, #MyResult);

  LastTimeSyncThis := pActTimeSyncElement^.pThis;
  TimeSyncTimeStamp := ops.tAbsolute;

END_FUNCTION

FUNCTION SafetyManager::TellAllInterfaceManagingModules
  VAR_INPUT
    pPara 	: ^CmdStruct;
    pResult 	: ^results;
    OverrideSync 	: BOOL;(* := FALSE *)
  END_VAR
  VAR
    pHelpManaging : ^t_ManagingComponent;
  END_VAR

  if pFirstManagingInterfaceComponent then
    pHelpManaging := pFirstManagingInterfaceComponent;
    while pHelpManaging do
      // call the newinst with the given parameters
      if pHelpManaging^.InfoBits.IsSynchron | OverrideSync then
        pHelpManaging^.pThis^.NewInst(pPara, pResult);
      end_if;

      pHelpManaging := pHelpManaging^.pNext;
    end_while;
  end_if;

END_FUNCTION

FUNCTION SafetyManager::SafetyManager
  VAR_OUTPUT
    ret_code 	: ConfStates;
  END_VAR
  VAR
    sd_retval : DINT;
  END_VAR

  //get interface for hardwaretree functions
  if ( OS_CILGET(INTERFACE_HARDWARETREE, #pHardwareTree)) then
    pHardwareTree := NIL;

    // logging can be used here already because the constructor of the base has been called before to initialize the log-interface-pointer
    LogError("@0457 (SafetyManager::SafetyManager) Hardwaretree-Interface not found. A newer OS is required for Safety-Modules");
  end_if;

  pTempMemCy := To_StdLib.Malloc(size:=SIZE_TEMP_MEMORY);
  if pTempMemCy then
    ud_SizeTempMemCy := SIZE_TEMP_MEMORY;
  else
    LogError("@0458 (SafetyManager::SafetyManager) Allocate temporary Memory failed");
  end_if;

  // try the new interface first
  sd_retval := OS_CILGet(INTERFACE_SAFETY_DLL2, #pSafetyDll2)$DINT;

  if sd_retval then
    // the new safety interface is not available => try the old one
    sd_retval := OS_CILGet(INTERFACE_SAFETY_DLL, #pSafetyDll)$DINT;

    if sd_retval then
      // no dll available
    elsif pSafetyDll^.version >= 5 then
      // dll available that allows quit error
      QuitErrorAvailable := 1;
    end_if;
  else
    // dll available that allows quit error and multiple connections
    QuitErrorAvailable := 2;
  end_if;

  OS_CILGet( INTERFACE_VARANMANAGER, #pVaran );

  ret_code := C_OK;

END_FUNCTION

FUNCTION SafetyManager::AllManagingNodesSynchron
  VAR_OUTPUT
    AllReady 	: BOOL;
  END_VAR
  VAR
    pHelpManaging : ^t_ManagingComponent;
    MyPara 	  : CmdStruct;
    MyResult	: results;
  END_VAR

  AllReady := TRUE;

  // check if any of the managing interface modules is not synchron
  if pFirstManagingInterfaceComponent then
    MyPara.uiCmd := CMD_SM_SYNC_CHECK;

    pHelpManaging := pFirstManagingInterfaceComponent;
    while pHelpManaging do
      // if any managing component isn't synchron => stop searching
      if pHelpManaging^.pThis^.NewInst(#MyPara, #MyResult) = ERROR then
        if (pHelpManaging^.InfoBits.IsOptional = TRUE) then
          if ((SafetyDomainTimeout & ((ops.tAbsolute - SynchroTimeout) > SafetyDomainTimeout))) then
            // we give up waiting => timeout exceeded
            b_SyncTimeoutExceeded := TRUE;
            // if it's the last managing module, then it's our connection to the master module
            if (IsTimeSyncMaster = 0) & pHelpManaging^.InfoBits.IsConnectionToMaster then
              // we have to be our own master now
              IsTimeSyncMaster := 1;
            end_if;
          else
            AllReady := FALSE;
          end_if;
        else
          AllReady := FALSE;
        end_if;

        // return; don't give up here => we have to check it for all domains, this one may be an optional interface frame domain
        pHelpManaging^.InfoBits.IsSynchron := FALSE;
      else
        pHelpManaging^.InfoBits.IsSynchron := TRUE;
      end_if;

      pHelpManaging := pHelpManaging^.pNext;
    end_while;
  end_if;

END_FUNCTION

FUNCTION SafetyManager::GetMasterConnection
  VAR_OUTPUT
    pMasterConn : ^t_ManagingComponent;
  END_VAR
  VAR
    pHelpManaging : ^t_ManagingComponent;
  END_VAR

  pMasterConn := NIL;

  if pFirstManagingInterfaceComponent then
    pHelpManaging := pFirstManagingInterfaceComponent;
    while pHelpManaging do
      if (pHelpManaging^.ModuleType = _VBC021Slave) | (pHelpManaging^.ModuleType = _VaranManager4VMC) | (pHelpManaging^.ModuleType = _GenericTimeSyncSlave) then
        pMasterConn := pHelpManaging;
        pMasterConn^.InfoBits.IsConnectionToMaster := TRUE;
        // if it's not the last in the list => we have to put it in the last place for easier timesync handling (last managing module to handle is the connection back to the master)
        if pMasterConn^.pNext then
          // if it's the first one
          if pMasterConn = pFirstManagingInterfaceComponent then
            pHelpManaging := pFirstManagingInterfaceComponent;
            while pHelpManaging^.pNext do
              pHelpManaging := pHelpManaging^.pNext;
            end_while;
            pFirstManagingInterfaceComponent := pFirstManagingInterfaceComponent^.pNext;
            pHelpManaging^.pNext := pMasterConn;
            pMasterConn^.pNext := NIL;
          else
            // if it's one in the middle
            pHelpManaging := pFirstManagingInterfaceComponent;
            while pHelpManaging^.pNext do
              if pHelpManaging^.pNext = pMasterConn then
                pHelpManaging^.pNext := pMasterConn^.pNext;
              end_if;

              pHelpManaging := pHelpManaging^.pNext;
            end_while;
            pHelpManaging^.pNext := pMasterConn;
            pMasterConn^.pNext := NIL;
          end_if;
        end_if;
        return;
      end_if;

      pHelpManaging := pHelpManaging^.pNext;
    end_while;
  end_if;

END_FUNCTION

FUNCTION SafetyManager::AddConfiguration
  VAR_INPUT
    Length 	: UINT;
    pData 	: ^void;
    IsFSoEConfig 	: BOOL;
  END_VAR
  VAR_OUTPUT
    retcode 	: DINT;
  END_VAR
  VAR
    pHelpCfg          : ^t_CfgListElem;
    pHelpModule       : ^t_ModuleListElem;
    pHelpPdo          : ^t_PdoListElem;
    pHelpSlave        : ^t_SlaveListElem;
    pHelpConnection   : ^t_FSoEConnectionDetails;
    pDataHelp         : ^void;
    i                 : UDINT;
    TmpPathLen        : UINT;
    TempCfgNo         : USINT;
    TempConnectionNo  : UINT;
    pHelpSafety       : ^t_SafetyComponent;
    pHelpManaging     : ^t_ManagingComponent;
    ModuleNo          : UDINT;
  END_VAR

(*
    Memory structure:
      4 Byte: SafetyNumber of CPU (is already there from initialisation in CSCP011_IM::InitSafeModule)
      1 Byte: Number of module configurations which are following
      for every module configuration (first is always the CPU itself)
        1 Byte: Info
        4 Byte: Interface Frame Source SafetyNumber (0 if it is no source for interface frames)
        4 Byte: Interface Frame CRC
        1 Byte: Number of destination inferface frame CRCs
        x Byte: Destination interface frame CRCs (number * sizeof(HDINT)
        2 Byte: Length of hardware path
        x Byte (depending on length in the 2 byte before): Hardwarepath
        2 Byte: Length of compressed hardware path
        x Byte (depending on length in the 2 byte before): Compressed Hardwarepath
        1 Byte: PDO out length for this module
      1 Byte: Number of pdo configurations which are following
      for every PDO configuration
        1 Byte: PDO length
        1 Byte: Interface frame info
        4 Byte: Interface CRC
        2 Byte: Length of source hardware path
        x Byte (depending on length in the 2 byte before): Hardwarepath of source
        2 Byte: Length of destination hardware path
        x Byte (depending on length in the 2 byte before): Hardwarepath of destination
      1 Byte: Number of slave configurations which are following
      for every slave configuration
        1 Byte: Info
        4 Byte: InterfaceCRC
        2 Byte: Length of hardware path
        x Byte (depending on length in the 2 byte before): Hardwarepath
        2 Byte: Length of compressed hardware path
        x Byte (depending on length in the 2 byte before): Compressed Hardwarepath

      if IsFSoEConfig = TRUE
      2 Byte: Number of connection infos which are following
      for every FSoE connection info
        2 Byte: ConnectionID
        1 Byte: ConnectionState
        1 Byte: Flags // Actually, type is 4 bytes in size but for compatibility reasons it is still used as 1 byte. As a result, bits 9-32 are currently not used.
        4 Byte: Master safety number

only if feature available:
        2 Byte: Transmission time in ms

        2 Byte: Offset where to read from master
        2 Byte: Size of data to read from master (and write to slave)
        2 Byte: Offset where to write to master
        2 Byte: Size of data to write to master (and read from slave)
        2 Byte: SlaveAddress
        2 Byte: Length of slave hardware path
        x Byte (depending on length in the 2 byte before): Slave hardware path
        2 Byte: Length of compressed slave hardware path
        x Byte (depending on length in the 2 byte before): Compressed slave hardware path
        2 Byte: Offset where to read from slave
        2 Byte: Offset where to write to slave

*)

  // check if the configuration is valid (pData <> NIL) & (Length must be at least 4 byte for SafetyNbr + 1 byte module cfg number + 1 byte pdo cfg number + 1 byte slave crc number)
  if pData & (Length >= 7)  then

    retcode := 0;

    // first we have to allocate some memory for the configuration
    if pConfigs = NIL then
      pConfigs$pVoid := To_StdLib.Malloc(size:=sizeof(t_CfgListElem));
      pHelpCfg := pConfigs;
    else
      pHelpCfg := pConfigs;
      while pHelpCfg^.pNext <> NIL do
        //if searched path is found, we already got this module in our list
        if pHelpCfg^.SafetyNbr = pData^$HDINT then
          // already in buffer => leave function
          return;
        else
          pHelpCfg := pHelpCfg^.pNext;
        end_if;
      end_while;

      //if searched path is found, we already got this module in our list
      if pHelpCfg^.SafetyNbr = pData^$HDINT then
        // already in buffer => leave function
        return;
      end_if;

      pHelpCfg^.pNext$pvoid := To_StdLib.Malloc(size:=sizeof(t_CfgListElem));
      pHelpCfg := pHelpCfg^.pNext;
    end_if;

    // if we have memory for the configuration => we add the data to the new element
    if pHelpCfg <> NIL then
      pDataHelp := pData;

      // set the next pointer to NIL
      pHelpCfg^.pNext := NIL;

      // safety number of the safety cpu
      pHelpCfg^.SafetyNbr := pDataHelp^$HDINT;
      pDataHelp += sizeof(HDINT);

      // number of module configurations which follow now
      TempCfgNo := pDataHelp^$USINT;
      pDataHelp += sizeof(USINT);

      pHelpCfg^.pFirstModuleCfg := NIL;

      // module configurations
      if TempCfgNo then
        for i := 0 to (TempCfgNo-1) do
          if pHelpCfg^.pFirstModuleCfg = NIL then
            pHelpCfg^.pFirstModuleCfg$pVoid := To_StdLib.Malloc(size:=sizeof(t_ModuleListElem));
            pHelpModule := pHelpCfg^.pFirstModuleCfg;
          else
            pHelpModule^.pNext$pvoid := To_StdLib.Malloc(size:=sizeof(t_ModuleListElem));
            pHelpModule := pHelpModule^.pNext;
          end_if;

          if pHelpModule then
            // initialize the pointers with NIL in case one of the mallocs fails
            pHelpModule^.ModuleInfo.pDestCRCs   := NIL;
            pHelpModule^.ModuleInfo.pPath       := NIL;
            pHelpModule^.ModuleInfo.pCompPath   := NIL;
            pHelpModule^.pNext                  := NIL;

            // info
            pHelpModule^.ModuleInfo.Info := pDataHelp^$BSINT;
            pDataHelp += sizeof(BSINT);

            // safety number of interface frame source
            pHelpModule^.ModuleInfo.SafetyNbr := pDataHelp^$HDINT;
            pDataHelp += sizeof(HDINT);

            // if it's the config owner => take the address service info to the info bits
            if pHelpCfg^.SafetyNbr = pHelpModule^.ModuleInfo.SafetyNbr then
              pHelpSafety := pFirstSafetyComponent;
              while pHelpSafety do
                // check if we got a component with this number
                if pHelpSafety^.SafetyNbr = pHelpCfg^.SafetyNbr then
                  pHelpSafety^.InfoBits.IsAddressService := pHelpModule^.ModuleInfo.Info.IsAddressService;
                end_if;

                pHelpSafety := pHelpSafety^.pNext;
              end_while;
            end_if;

            // interface CRC of interface frame
            pHelpModule^.ModuleInfo.InterfaceCRC := pDataHelp^$HDINT;
            pDataHelp += sizeof(HDINT);

            if pHelpModule^.ModuleInfo.InterfaceCRC then
              // someone might connect to us via udp because we supply an interface frame
              sUdpVars.UdpInit.ProvidesIF := TRUE;
            end_if;

            // interface frame destination CRCs
            if pHelpModule^.ModuleInfo.Info.IsInterfaceDest then
              // number of CRCs
              TmpPathLen := pDataHelp^$USINT; // save some time with this local variable
              pHelpModule^.ModuleInfo.DestCRCNo := TmpPathLen$USINT;
              pDataHelp += sizeof(USINT);

              // allocate memory for the module path
              pHelpModule^.ModuleInfo.pDestCRCs$pVoid := To_StdLib.Malloc(size:=TmpPathLen * sizeof(HDINT));
              if pHelpModule^.ModuleInfo.pDestCRCs = NIL then
                ClassState := -1;
                retcode := -2;
                return;
              end_if;

              // save CRCs
              _memcpy(ptr1:=pHelpModule^.ModuleInfo.pDestCRCs, ptr2:=pDataHelp, cntr:=TmpPathLen * sizeof(HDINT));
              pDataHelp += TmpPathLen * sizeof(HDINT);
            else
              pHelpModule^.ModuleInfo.DestCRCNo := 0;
              pHelpModule^.ModuleInfo.pDestCRCs := NIL;
            end_if;

            // length of hardwarepath
            TmpPathLen := pDataHelp^$UINT; // save some time with this local variable
            pHelpModule^.ModuleInfo.PathLen := TmpPathLen;
            pDataHelp += sizeof(UINT);

            // allocate memory for the module path
            pHelpModule^.ModuleInfo.pPath$pVoid := To_StdLib.Malloc(size:=TmpPathLen);
            if pHelpModule^.ModuleInfo.pPath = NIL then
              ClassState := -1;
              retcode := -2;
              return;
            end_if;

            // save hardwarepath
            _memcpy(ptr1:=pHelpModule^.ModuleInfo.pPath, ptr2:=pDataHelp, cntr:=TmpPathLen);
            pDataHelp += TmpPathLen;

            // length of hardwarepath
            TmpPathLen := pDataHelp^$UINT; // save some time with this local variable
            pHelpModule^.ModuleInfo.CompPathLen := TmpPathLen;
            pDataHelp += sizeof(UINT);

            // allocate memory for the module path
            pHelpModule^.ModuleInfo.pCompPath$pVoid := To_StdLib.Malloc(size:=TmpPathLen);
            if pHelpModule^.ModuleInfo.pCompPath = NIL then
              ClassState := -1;
              retcode := -2;
              return;
            end_if;

            // save compressed hardwarepath
            _memcpy(ptr1:=pHelpModule^.ModuleInfo.pCompPath, ptr2:=pDataHelp, cntr:=TmpPathLen);
            pDataHelp += TmpPathLen;

            // PDO out length for this module (to assign the length to the pdo configurations)
            pHelpModule^.ModuleInfo.PdoOutLen := pDataHelp^$USINT;
            pDataHelp += sizeof(USINT);
          else
            ClassState := -1;
            retcode := -2;
            return;
          end_if;
        end_for;
      end_if;

      // number of Pdo configurations which follow now
      TempCfgNo := pDataHelp^$USINT;
      pDataHelp += sizeof(USINT);

      pHelpCfg^.pFirstPdoCfg := NIL;

      // Pdo configurations
      if TempCfgNo then
        for i := 0 to (TempCfgNo-1) do
          if pHelpCfg^.pFirstPdoCfg = NIL then
            pHelpCfg^.pFirstPdoCfg$pVoid := To_StdLib.Malloc(size:=sizeof(t_PdoListElem));
            pHelpPdo := pHelpCfg^.pFirstPdoCfg;
          else
            pHelpPdo^.pNext$pvoid := To_StdLib.Malloc(size:=sizeof(t_PdoListElem));
            pHelpPdo := pHelpPdo^.pNext;
          end_if;

          if pHelpPdo then
            // initialize the pointers with NIL in case one of the mallocs fails
            pHelpPdo^.PdoInfo.pSourcePath     := NIL;
            pHelpPdo^.PdoInfo.pDestPath       := NIL;
            pHelpPdo^.pNext                   := NIL;

            // pdo length
            pHelpPdo^.PdoInfo.PdoLen := pDataHelp^$USINT;
            pDataHelp += sizeof(USINT);

            // is it an interface pdo?
            pHelpPdo^.PdoInfo.Info := pDataHelp^$BSINT;
            pDataHelp += sizeof(BSINT);

            // if it is an interface frame, we have to copy the CRC too
            if pHelpPdo^.PdoInfo.Info.IsInterfacePDO then
              // interface CRC
              pHelpPdo^.PdoInfo.InterfaceCRC := pDataHelp^$HDINT;
            else
              pHelpPdo^.PdoInfo.InterfaceCRC := 0;
            end_if;
            pDataHelp += sizeof(HDINT);

            // length of source hardwarepath
            TmpPathLen := pDataHelp^$UINT; // save some time with this local variable
            pHelpPdo^.PdoInfo.SourcePathLen := TmpPathLen;
            pDataHelp += sizeof(UINT);

            // allocate memory for the source module path
            pHelpPdo^.PdoInfo.pSourcePath$pVoid := To_StdLib.Malloc(size:=TmpPathLen);
            if pHelpPdo^.PdoInfo.pSourcePath = NIL then
              ClassState := -1;
              retcode := -2;
              return;
            end_if;

            // save source hardwarepath
            _memcpy(ptr1:=pHelpPdo^.PdoInfo.pSourcePath, ptr2:=pDataHelp, cntr:=TmpPathLen);
            pDataHelp += TmpPathLen;

            // check for an IP Address
            if pHelpPdo^.PdoInfo.Info.SrcPathIsCompressed & (pHelpPdo^.PdoInfo.pSourcePath^$USINT = INTERFACE_IP_MODE) then
              // add the connection (we're consumer and we got the IP address of the producer)
              AddUdpConnection(IP:=(pHelpPdo^.PdoInfo.pSourcePath$^HDINT + 5)^, IFCRC:=(pHelpPdo^.PdoInfo.pSourcePath$^HDINT + 1)^, SafetyNumber:=pHelpCfg^.SafetyNbr, ProducerList:=TRUE);
            end_if;

            // length of destination hardwarepath
            TmpPathLen := pDataHelp^$UINT; // save some time with this local variable
            pHelpPdo^.PdoInfo.DestPathLen := TmpPathLen;
            pDataHelp += sizeof(UINT);

            // allocate memory for the destination module path
            pHelpPdo^.PdoInfo.pDestPath$pVoid := To_StdLib.Malloc(size:=TmpPathLen);
            if pHelpPdo^.PdoInfo.pDestPath = NIL then
              ClassState := -1;
              retcode := -2;
              return;
            end_if;

            // save destination hardwarepath
            _memcpy(ptr1:=pHelpPdo^.PdoInfo.pDestPath, ptr2:=pDataHelp, cntr:=TmpPathLen);
            pDataHelp += TmpPathLen;

            // check if a prior configuration also added this PDO (possible if a CSTO gets PDOs from 2 CSCPs)
            if DoublePDOEntry(pHelpPdo^.PdoInfo, pHelpCfg) then
              // use ID 255 (as kind of invalid) and mark the PDO as double entry (will not be distributed then)
              pHelpPdo^.PdoInfo.PDO_ID := 255;
              pHelpPdo^.PdoInfo.Info.DoublePDOEntry := TRUE;
            else
              // now we give it a priority and increase the number for the next pdo
              pHelpPdo^.PdoInfo.PDO_ID := ActPDO_ID;
              ActPDO_ID += 1;
            end_if;

          else
            ClassState := -1;
            retcode := -2;
            return;
          end_if;
        end_for;
      end_if;

      // number of slave configurations which follow now
      TempCfgNo := pDataHelp^$USINT;
      pDataHelp += sizeof(USINT);

      pHelpCfg^.pFirstSlaveCfg:= NIL;

      // slave configurations
      if TempCfgNo then
        for i := 0 to (TempCfgNo-1) do
          if pHelpCfg^.pFirstSlaveCfg = NIL then
            pHelpCfg^.pFirstSlaveCfg$pVoid := To_StdLib.Malloc(size:=sizeof(t_SlaveListElem));
            pHelpSlave := pHelpCfg^.pFirstSlaveCfg;
          else
            pHelpSlave^.pNext$pvoid := To_StdLib.Malloc(size:=sizeof(t_SlaveListElem));
            pHelpSlave := pHelpSlave^.pNext;
          end_if;

          if pHelpSlave then
            // initialize the pointers with NIL in case one of the mallocs fails
            pHelpSlave^.SlaveInfo.pPath     := NIL;
            pHelpSlave^.SlaveInfo.pCompPath := NIL;
            pHelpSlave^.pNext               := NIL;

            // info
            pHelpSlave^.SlaveInfo.Info := pDataHelp^$BSINT;
            pDataHelp += sizeof(BSINT);

            // InterfaceCRC
            pHelpSlave^.SlaveInfo.InterfaceCRC := pDataHelp^$HDINT;
            pDataHelp += sizeof(HDINT);

            // length of hardwarepath
            TmpPathLen := pDataHelp^$UINT; // save some time with this local variable
            pHelpSlave^.SlaveInfo.PathLen := TmpPathLen;
            pDataHelp += sizeof(UINT);

            // allocate memory for the module path
            pHelpSlave^.SlaveInfo.pPath$pVoid := To_StdLib.Malloc(size:=TmpPathLen);
            if pHelpSlave^.SlaveInfo.pPath = NIL then
              ClassState := -1;
              retcode := -2;
              return;
            end_if;

            // save hardwarepath
            _memcpy(ptr1:=pHelpSlave^.SlaveInfo.pPath, ptr2:=pDataHelp, cntr:=TmpPathLen);
            pDataHelp += TmpPathLen;

            // length of hardwarepath
            TmpPathLen := pDataHelp^$UINT; // save some time with this local variable
            pHelpSlave^.SlaveInfo.CompPathLen := TmpPathLen;
            pDataHelp += sizeof(UINT);

            // allocate memory for the module path
            pHelpSlave^.SlaveInfo.pCompPath$pVoid := To_StdLib.Malloc(size:=TmpPathLen);
            if pHelpSlave^.SlaveInfo.pCompPath = NIL then
              ClassState := -1;
              retcode := -2;
              return;
            end_if;

            // save compressed hardwarepath
            _memcpy(ptr1:=pHelpSlave^.SlaveInfo.pCompPath, ptr2:=pDataHelp, cntr:=TmpPathLen);
            pDataHelp += TmpPathLen;
          else
            ClassState := -1;
            retcode := -2;
            return;
          end_if;
        end_for;
      end_if;

      pHelpCfg^.pFirstFSoEConnection := NIL;

      // check if it's a FSoE Config
      if IsFSoEConfig then
        // number of connection details which follow now
        TempConnectionNo := pDataHelp^$UINT;
        pDataHelp += sizeof(UINT);

        // if we got connections
        if TempConnectionNo then
          for i := 0 to (TempConnectionNo-1) do
            if pHelpCfg^.pFirstFSoEConnection = NIL then
              pHelpCfg^.pFirstFSoEConnection$pVoid := To_StdLib.Malloc(size:=sizeof(t_FSoEConnectionDetails));
              pHelpConnection := pHelpCfg^.pFirstFSoEConnection;
            else
              pHelpConnection^.pNext$pvoid := To_StdLib.Malloc(size:=sizeof(t_FSoEConnectionDetails));
              pHelpConnection := pHelpConnection^.pNext;
            end_if;

            // if we succeeded to allocate memory
            if pHelpConnection then
              // initialize the pointers with NIL in case one of the mallocs fails
              pHelpConnection^.pSlavePath       := NIL;
              pHelpConnection^.pSlavePathComp   := NIL;
              pHelpConnection^.pNext            := NIL;
              pHelpConnection^.pNextSorted      := NIL;

              // connection ID
              pHelpConnection^.ConnectionID := pDataHelp^$UINT;
              pDataHelp += sizeof(UINT);

              // connection state (use our own state internally)
              pHelpConnection^.InternalConnectionState := FCS_RESET;
              pHelpConnection^.ConnectionState := pDataHelp^$t_FSoEConnectionState;

              pDataHelp += sizeof(USINT);

              // flags

              // Actually, type is 4 bytes in size but for compatibility reasons it is still used as 1 byte. As a result, bits 9-32 are currently not used.
              if bdFeatureEnable.FSoEFlags_4ByteSize then
                pHelpConnection^.Flags$t_FSoEFlags := pDataHelp^$t_FSoEFlags;
                pDataHelp += sizeof(t_FSoEFlags);
              else
                pHelpConnection^.Flags$USINT := pDataHelp^$USINT;
                pDataHelp += sizeof(USINT);
              end_if;

              // check if FlexCon functionality is used according to the flags in this connection
              if (pHelpConnection^.Flags AND SM_FLAGS_FLEXCON_MASK) = SM_FLAGS_FLEXCON_HOST then
                // if there are no generic dynamic FSoE devices registered (this is to prevent the FlexCon functionality from conflicting with the MultiModule used for the LogiMover)
                if GetModuleTypeNo(ModuleType:=_GenericDynamicFSoE) = 0 then
                  if sFlexCon.Role = _FlexConNode then
                    sFlexCon.Role := _InvalidConstellation;
                  elsif sFlexCon.Role <> _InvalidConstellation then
                    sFlexCon.Role := _FlexConHost;

                    pHelpSafety := pFirstSafetyComponent;
                    while pHelpSafety do
                      // check if we got an address service
                      if pHelpSafety^.InfoBits.IsAddressService then
                        // check if it's NIL or already our desired value
                        if (sFlexCon.pSafetyHost = NIL) | (sFlexCon.pSafetyHost = pHelpSafety) then
                          // remember the pointer for quick access later
                          sFlexCon.pSafetyHost := pHelpSafety;
                        else
                          LogError(e_msg:="@05DA (SafetyManager::AddConfiguration) Multiple FlexConHosts found! Check Safety Designer Projects of all connected Safe CPUs");

                          sFlexCon.Role := _InvalidConstellation;
                        end_if;
                      end_if;

                      pHelpSafety := pHelpSafety^.pNext;
                    end_while;
                  end_if;
                end_if;
              elsif (pHelpConnection^.Flags AND SM_FLAGS_FLEXCON_MASK) = SM_FLAGS_FLEXCON_NODE then
#ifdef SAFETY_DEBUG_LOGGING_ACTIVATED
                LogError(e_msg:="@DBG SafetyManager: Found FSOE Connection of FlexConNode");

                LogValue(pString:="Number of VBC021_Slave objects with safety memory: 0x{0}", Value:=GetModuleTypeNo(ModuleType:=_VBC021Slave));
                LogValue(pString:="Number of VM objects with safety memory: 0x{0}", Value:=GetModuleTypeNo(ModuleType:=_VaranManager4VMC));
#endif
                // if we detected a Node but the role has already been set to Host
                if sFlexCon.Role = _FlexConHost then
                  // it's an invalid constellation (can't be host and node at the same time)
                  sFlexCon.Role := _InvalidConstellation;
                elsif sFlexCon.Role <> _InvalidConstellation then

                  // check if there is only one possible connection to the host
                  ModuleNo := GetModuleTypeNo(ModuleType:=_VBC021Slave) + GetModuleTypeNo(ModuleType:=_VaranManager4VMC);
                  if ModuleNo = 1 then
                    sFlexCon.Role := _FlexConNode;

                    // get the managing module connecting us with the host
                    pHelpManaging := pFirstManagingInterfaceComponent;
                    while pHelpManaging do
                      if (pHelpManaging^.ModuleType = _VBC021Slave) | (pHelpManaging^.ModuleType = _VaranManager4VMC) then
                        // remember the pointer for quick access later
                        sFlexCon.pManaging2Host := pHelpManaging;
                      end_if;

                      pHelpManaging := pHelpManaging^.pNext;
                    end_while;
                  else
                    // invalid
                    sFlexCon.Role := _InvalidConstellation;

                    // check if there are no or too many vbc021 slave modules
                    if ModuleNo = 0 then
                      LogError(e_msg:="@05DB (SafetyManager::AddConfiguration) No VBC021_Slave with defined safety memory detected");
                    else
                      LogError(e_msg:="@05DD (SafetyManager::AddConfiguration) More than 1 VBC021_Slave detected => NOT ALLOWED!");
                    end_if;
                  end_if;
                end_if;
              end_if;

              // master safety number
              pHelpConnection^.OwnerSafetyNbr := pDataHelp^$HDINT;
              pDataHelp += sizeof(HDINT);

              // the feature is not available in older safety module classes, so we have to do this for compatibility reasons
              if bdFeatureEnable.TransmissionTimeInConfig then
                // transmission time in ms
                pHelpConnection^.TransmissionTime_ms := pDataHelp^$UINT;
                pDataHelp += sizeof(UINT);
              else
                pHelpConnection^.TransmissionTime_ms := 0;
              end_if;

              // offset where to read from master
              pHelpConnection^.MasterReadOffset := pDataHelp^$UINT;
              pDataHelp += sizeof(UINT);

              // size of data to read from master (and write to slave)
              pHelpConnection^.MasterReadSize := pDataHelp^$UINT;
              pDataHelp += sizeof(UINT);

              // offset where to write to master
              pHelpConnection^.MasterWriteOffset := pDataHelp^$UINT;
              pDataHelp += sizeof(UINT);

              // size of data to write to master (and read from slave)
              pHelpConnection^.MasterWriteSize := pDataHelp^$UINT;
              pDataHelp += sizeof(UINT);

              // slave address
              pHelpConnection^.SlaveAddress := pDataHelp^$UINT;
              pDataHelp += sizeof(UINT);

              // wait for slave addresses if any connection is not initialized
              if (pHelpConnection^.ConnectionState = FCS_NOT_INITIALIZED) & (pHelpConnection^.SlaveAddress = 0) then
                b_AllLocalSlaveAddressesValid := FALSE;
              end_if;

              // length of uncompressed slave hardwarepath
              TmpPathLen := pDataHelp^$UINT; // save some time with this local variable
              pHelpConnection^.SlavePathLen := TmpPathLen;
              pDataHelp += sizeof(UINT);

              if pHelpConnection^.Flags.IsMaster then
                // allocate memory for the module path
                pHelpConnection^.pSlavePath$pVoid := To_StdLib.Malloc(size:=TmpPathLen);
                if pHelpConnection^.pSlavePath = NIL then
                  ClassState := -1;
                  retcode := -2;
                  return;
                end_if;

                // save hardwarepath
                _memcpy(ptr1:=pHelpConnection^.pSlavePath, ptr2:=pDataHelp, cntr:=TmpPathLen);
                pDataHelp += TmpPathLen;
              end_if;

              // length of compressed slave hardwarepath
              TmpPathLen := pDataHelp^$UINT; // save some time with this local variable
              pHelpConnection^.SlavePathCompLen := TmpPathLen;
              pDataHelp += sizeof(UINT);

              if pHelpConnection^.Flags.IsMaster then
                // allocate memory for the module path
                pHelpConnection^.pSlavePathComp$pVoid := To_StdLib.Malloc(size:=TmpPathLen);
                if pHelpConnection^.pSlavePathComp = NIL then
                  ClassState := -1;
                  retcode := -2;
                  return;
                end_if;

                // save compressed hardwarepath
                _memcpy(ptr1:=pHelpConnection^.pSlavePathComp, ptr2:=pDataHelp, cntr:=TmpPathLen);
                pDataHelp += TmpPathLen;

                // if it's a udp connection, consider the transmission time
                if (pHelpConnection^.pSlavePathComp^ = INTERFACE_IP_MODE) & pHelpConnection^.TransmissionTime_ms then
                  if pHelpConnection^.TransmissionTime_ms < sUdpVars.LowestTransmissionTime_ms then
                    sUdpVars.LowestTransmissionTime_ms := pHelpConnection^.TransmissionTime_ms;
                  end_if;
                end_if;
              end_if;

              // offset where to read from master
              pHelpConnection^.SlaveReadOffset := pDataHelp^$UINT;
              pDataHelp += sizeof(UINT);

              // offset where to write to master
              pHelpConnection^.SlaveWriteOffset := pDataHelp^$UINT;
              pDataHelp += sizeof(UINT);

              // initialize log marker
              pHelpConnection^.bsLogError := 0;
            else
              ClassState := -1;
              retcode := -2;
              return;
            end_if;
          end_for;
        end_if;
      end_if;

      ConfigNo += 1;

      // check if the given size matches the memory structure
      if (pDataHelp$UDINT - pData$UDINT) <> Length then
        LogError("@0459 (SafetyManager::AddConfiguration) Invalid configuration data given (length doesn't match memory structure)");
        retcode := -3;
        return;
      end_if;
    else
      ClassState := -1;
      retcode := -2;
      return;
    end_if;
  else
    // invalid configuration
    LogError("@045A (SafetyManager::AddConfiguration) Found invalid safety cpu configuration: Pointer or size wrong");
    retcode := -1;
  end_if;

END_FUNCTION

FUNCTION SafetyManager::FreeCfgLists
  VAR
    pHelpCfg        : ^t_CfgListElem;
    pHelpModule     : ^t_ModuleListElem;
    pHelpPdo        : ^t_PdoListElem;
    pHelpConnection : ^t_FSoEConnectionDetails;
  END_VAR

  while pConfigs do
    pHelpCfg := pConfigs;
    pConfigs := pConfigs^.pNext;

    // while we got module cfgs
    while pHelpCfg^.pFirstModuleCfg do
      pHelpModule := pHelpCfg^.pFirstModuleCfg;
      pHelpCfg^.pFirstModuleCfg := pHelpCfg^.pFirstModuleCfg^.pNext;

      if pHelpModule^.ModuleInfo.pDestCRCs then
        To_StdLib.Free(pHelpModule^.ModuleInfo.pDestCRCs);
      end_if;

      To_StdLib.Free(pHelpModule^.ModuleInfo.pPath);
      To_StdLib.Free(pHelpModule^.ModuleInfo.pCompPath);
      To_StdLib.Free(pHelpModule);
    end_while;

    // while we got pdo cfgs
    while pHelpCfg^.pFirstPdoCfg do
      pHelpPdo := pHelpCfg^.pFirstPdoCfg;
      pHelpCfg^.pFirstPdoCfg := pHelpCfg^.pFirstPdoCfg^.pNext;

      To_StdLib.Free(pHelpPdo^.PdoInfo.pSourcePath);
      To_StdLib.Free(pHelpPdo^.PdoInfo.pDestPath);
      To_StdLib.Free(pHelpPdo);
    end_while;

    // while we got connection infos
    while pHelpCfg^.pFirstFSoEConnection do
      pHelpConnection := pHelpCfg^.pFirstFSoEConnection;
      pHelpCfg^.pFirstFSoEConnection := pHelpCfg^.pFirstFSoEConnection^.pNext;

      if pHelpConnection^.pSlavePath then
        To_StdLib.Free(mptr:=pHelpConnection^.pSlavePath);
      end_if;

      if pHelpConnection^.pSlavePathComp then
        To_StdLib.Free(mptr:=pHelpConnection^.pSlavePathComp);
      end_if;

      To_StdLib.Free(mptr:=pHelpConnection);
    end_while;

    To_StdLib.Free(pHelpCfg);
  end_while;
  pSortedConnections := NIL; // may have contained a pointer within the config (to the connection with the lowest slave address)
  ConfigNo := 0;

END_FUNCTION

FUNCTION SafetyManager::AddOwnCPUsToList
  VAR
    pHelpSafety : ^t_SafetyComponent;
  END_VAR

  // reset number of memorized safe cpu numbers
  SafeCPU_Nbr_No := 0;

  // check if any of the managing modules is not synchron
  if pFirstSafetyComponent then
    pHelpSafety := pFirstSafetyComponent;
    while pHelpSafety do
      // add all safety cpus to the parameters
      if IsCPUModule(pHelpSafety^.ModuleType) then
        if pHelpSafety^.SafetyNbr then
          aSafetyCPU_Nbr[SafeCPU_Nbr_No] := pHelpSafety^.SafetyNbr;
          SafeCPU_Nbr_No += 1;
        end_if;
      end_if;

      pHelpSafety := pHelpSafety^.pNext;
    end_while;
  end_if;

END_FUNCTION

FUNCTION SafetyManager::AllCPUConfigsArrived
  VAR_OUTPUT
    AllReady 	: BOOL;
  END_VAR
  VAR
    pHelpCfg : ^t_CfgListElem;
    i : UDINT;
    Found : BOOL;
  END_VAR

  // check if there are any CPUs
  if SafeCPU_Nbr_No then
    // if we have already all configurations (according to the number) check if they are correct
    if ConfigNo = SafeCPU_Nbr_No then

      // normally we should be fine now
      AllReady := TRUE;

      // check all safety numbers stored
      for i := 0 to SafeCPU_Nbr_No-1 do

        Found := FALSE;

        // search all configurations
        pHelpCfg := pConfigs;
        while pHelpCfg do
          // if we found a match => stop searching for this one
          if pHelpCfg^.SafetyNbr = aSafetyCPU_Nbr[i] then
            Found := TRUE;
            exit;
          end_if;
          pHelpCfg := pHelpCfg^.pNext;
        end_while;

        // if this configuration hasn't been found, we may have a problem
        if Found = FALSE then
          AllReady := FALSE;
          LogError("@045B (SafetyManager::AllCPUConfigsArrived) Invalid CPU configuration found!");
          return;
        end_if;
      end_for;
    else
      AllReady := FALSE;

      if ConfigNo > SafeCPU_Nbr_No then
        LogError("@045C (SafetyManager::AllCPUConfigsArrived) ERROR! More configs available than safety CPUs");
      end_if;
    end_if;
  else
    AllReady := TRUE;
    LogError("@045D (SafetyManager::AllCPUConfigsArrived) No Safety CPU found in the system!");
  end_if;

END_FUNCTION

FUNCTION SafetyManager::AddLocalCPUCfg
  VAR_INPUT
    Length 	: UINT;
    pData 	: ^void;
    IsFSoECfg 	: BOOL;(* := FALSE *)
  END_VAR
  VAR
    pHelpLocalCfg   : ^t_LocalCfgListElem;
    EditOldCfg      : BOOL;
  END_VAR

  LastCfgReceiveTime := ops.tAbsolute;

  // if the a module wants to add the config which is already added => overwrite the old config
  EditOldCfg := FALSE;

  if pFirstLocalCPUCfg = NIL then
    pFirstLocalCPUCfg$pVoid := To_StdLib.Malloc(size:=sizeof(t_LocalCfgListElem));
    pHelpLocalCfg := pFirstLocalCPUCfg;
  else
    pHelpLocalCfg := pFirstLocalCPUCfg;

    if pHelpLocalCfg^.SafetyNbr = pData^$HDINT then
      EditOldCfg := TRUE;
    else
      while pHelpLocalCfg^.pNext <> NIL do
        pHelpLocalCfg := pHelpLocalCfg^.pNext;
        if pHelpLocalCfg^.SafetyNbr = pData^$HDINT then
          EditOldCfg := TRUE;
          exit;
        end_if;
      end_while;
      if EditOldCfg = FALSE then
        pHelpLocalCfg^.pNext$pVoid := To_StdLib.Malloc(size:=sizeof(t_LocalCfgListElem));

        pHelpLocalCfg := pHelpLocalCfg^.pNext;
      end_if;
    end_if;
  end_if;

  if pHelpLocalCfg <> NIL then
    pHelpLocalCfg^.SafetyNbr          := pData^$HDINT;
    pHelpLocalCfg^.ConfigSize         := Length;
    pHelpLocalCfg^.pConfig            := pData;  // memory can be accessed always (never freed)
    pHelpLocalCfg^.ConfigSent2Master  := FALSE;
    pHelpLocalCfg^.IsFSoECfg          := IsFSoECfg;

    if IsFSoECfg then
      sUdpVars.UdpInit.FSoEAvailable := TRUE;
    end_if;

    // only if we created a new element (incrementing has to be done last because of thread safety: bg increments the value and cyclic uses the list)
    if EditOldCfg = FALSE then
      pHelpLocalCfg^.pNext := NIL;
      LocalCPUCfgNo += 1;

      // new cpu config => reinitalize everything
      ReinitEverything();
    end_if;
  else
    ClassState := -1;
    LogError("@045E (SafetyManager::AddLocalCPUCfg) Failed to allocate Memory for the local CPU Configuration");
  end_if;

END_FUNCTION

FUNCTION SafetyManager::SendLocalCfgsToMaster
  VAR
    pHelpLocalCfg : ^t_LocalCfgListElem;
    i : UDINT;
  END_VAR

  if LocalCPUCfgNo then
    pHelpLocalCfg := pFirstLocalCPUCfg;

    for i := 0 to (LocalCPUCfgNo-1) do
      if pHelpLocalCfg^.ConfigSize then
        // if we're the master, we keep the configuration of this cpu and share the essentials later (when we got all configurations) with all other domains (distribute the mapping)
        if AddConfiguration(pHelpLocalCfg^.ConfigSize, pHelpLocalCfg^.pConfig, pHelpLocalCfg^.IsFSoECfg) <> 0 then
          LogError("@045F (SafetyManager::SendLocalCfgsToMaster) Failed to add a safety cpu configuration to the local config-memory");
        end_if;
      end_if;

      pHelpLocalCfg := pHelpLocalCfg^.pNext;
    end_for;
  end_if;

END_FUNCTION

FUNCTION SafetyManager::BroadCastActPDO
  VAR
    MyPara 	  : CmdStruct;
    PdoMemSize : UINT;
    pPdoMem    : ^USINT;
    pHelp      : ^USINT;
    TmpPathLen : UINT;
    SourceDest : t_SourceDest;
    SafetyNbr           : HDINT;
  END_VAR

  // put pdo (marked by pActualSendPDO) into linear memory, find out who needs it and broadcast it

(*
    Memory structure:
      1 Byte: Number of Domains involved
      x Byte: 1 Byte for every involved Domain number
      1 Byte: Number of Domains in source path
      x Byte: 1 Byte for every domain in source path
      1 Byte: Number of Domains in destination path
      x Byte: 1 Byte for every domain in destination path
      1 Byte: ID of this PDO (starting at 0)
      1 Byte: Length of PDO
      1 Byte: Is it an interface frame
      4 Byte: Interface CRC
      2 Byte: Length of source hardware path
      x Byte (depending on length in the 2 byte before): Hardwarepath of source
      2 Byte: Length of destination hardware path
      x Byte (depending on length in the 2 byte before): Hardwarepath of destination
*)

  // if the pointer is NIL or it's an interface frame broadcast, don't distribute it, there are virtual PDOs to be distributed instead of the broadcasts (if necessary)
  if (pActualSendPDO = NIL) | pActualSendPDO^.PdoInfo.Info.IFBroadCast then
    return;
  end_if;

  // add up the sizes and allocate the memory
  PdoMemSize := sizeof(USINT) +                           // 1 byte number of domains involved
                1 +                                       // 1 byte for every involved domain
                sizeof(USINT) +                           // 1 byte number of domains in source path
                1 +                                       // 1 byte for every domain in source path
                sizeof(USINT) +                           // 1 byte number of domains in destination path
                1 +                                       // 1 byte for every domain in destination path
                sizeof(USINT) +                           // 1 byte ID of this PDO (starting at 0)
                sizeof(USINT) +                           // 1 byte length of PDO
                sizeof(t_PdoCfgInfo) +                    // 1 byte pdo info (is it interface frame or optional...)
                sizeof(HDINT) +                           // 4 byte interface CRC
                sizeof(UINT) +                            // 2 byte length of source hardware path
                pActualSendPDO^.PdoInfo.SourcePathLen +   // x byte source hardware path
                sizeof(UINT) +                            // 2 byte length of destination hardware path
                pActualSendPDO^.PdoInfo.DestPathLen;      // x byte destination hardware path
